FUNCTION_BLOCK FB_Conveyor
VAR_INPUT
	bEnable	: BOOL;
END_VAR
VAR_OUTPUT
	bRunning	: BOOL;
END_VAR
VAR
	fSpeed		: LREAL;
	bStartReq	: BOOL;
END_VAR

bRunning := bEnable AND bStartReq AND fSpeed > 0;

PROPERTY Speed : LREAL
GET // PUBLIC
Speed := fSpeed;
END_GET
SET // PUBLIC
fSpeed := F_Clamp(Speed, 0, GVL_Parameters.fMaxSpeed);
END_SET
END_PROPERTY

METHOD Start : BOOL
bStartReq := bEnable;
Start := bStartReq;
END_METHOD

METHOD Stop
bStartReq := FALSE;
END_METHOD

END_FUNCTION_BLOCK

(* stored: Version 1.1.0.1
   POU FB_Conveyor: Id {c67dcc1c-41b3-4dfe-9469-81846a2ee30b}, SpecialFunc None
   Property Speed: Id {7f5b5d05-382f-434b-9a3f-d61a6b8f8231}
   Get Get: Id {4b3dfed5-05d7-46e6-b145-445085d51ba8}
   Set Set: Id {a864b4f8-ba8f-4f6f-ad8c-12e35bac562a}
   Method Start: Id {1b3e6602-7884-4fb4-b326-99630cc286c9}
   Method Stop: Id {713dbbbc-37e5-4f78-9aad-2cff70743fac} *)
